Staubli VAL3: HMI_safezone.pjx

--- HMI_safezone.pjx ---
Parameters version=s8.15Cs9_BS3113 stackSize=5000 millimeterUnit=true
Program file=bind.pgx
Program file=main.pgx
Program file=movePoint.pgx
Program file=onStart.pgx
Program file=refreshData.pgx
Program file=setData.pgx
Program file=setFrameData.pgx
Program file=start.pgx
Program file=stop.pgx
Program file=teachPoint.pgx
Data file=HMI_safezone.dtx
Library alias=safeTemp path=Disk://data/CustomerLib/default/safeData/safeData.pjx
Library alias=util path=Disk://HMI_cs9/HMI_util/HMI_util.pjx
Library alias=safeCheck path=Disk://source/projectSource/safeCheck/safeCheck.pjx
Library alias=saveData path=Disk://source/saveData/saveData.pjx

--- HMI_safezone.dtx ---
mdesc mNomSpeed = {blend=off}
string sList
string sSelZone
bool bSetFrame
bool bTeach1
bool bMove
bool bRename
bool bConfirm
bool bActive
public num nFrame[6]
num nTRSF1[6]
num nTRSF2[6]
string sLastZone
num _nZoneIndex
string sComment
frame fFrame = {fatherId=world[0]}
bool bBack
tool tTool = {fatherId=flange[0]}
bool bSetFrameData
string sToolIndex

--- main.pgx ---
public program main()
  local bool l_bResult
  local bool l_bExit
begin
  do
    if util:sPage!="safezone"
      util:sPage="safezone"
      call util:loadingPage()
      call onStart()
      call bind()
      userPage(util:sPage)
      delay(0.5)
    endIf

    if sSelZone!=sLastZone and sSelZone!=""
      sLastZone=sSelZone
      toNum(sLastZone,_nZoneIndex,l_bResult)
      bActive=(safeTemp:zZoneItem[_nZoneIndex].bActive==true)
      call refreshData(_nZoneIndex)
    endIf
    if bSetFrame
      //      util:sPage="Wizard"
      //      userPage(util:sPage)
      bSetFrame=false
      //      popUpMsg("设定坐标系")
      //      call refreshData(_nZoneIndex)
    elseIf bSetFrameData
      bSetFrameData=false
      call setFrameData(_nZoneIndex)
      call refreshData(_nZoneIndex)

    elseIf bTeach1
      bTeach1=false
      call teachPoint(_nZoneIndex)
      call refreshData(_nZoneIndex)
    elseIf bMove
      bMove=false
      call movePoint(_nZoneIndex)
    elseIf bConfirm
      bConfirm=false
      call setData(_nZoneIndex)
      call refreshData(_nZoneIndex)
    elseIf bBack
      bBack=false
      l_bExit=true
    endIf

    delay(0)
  until l_bExit==true
  call saveData:setBaseJOG(saveData:nJogTool)
end

--- start.pgx ---
program start()
begin
end

--- bind.pgx ---
program bind()
  local string l_nmb
  local num l_i
begin
  userPageBindClick("safezone","btnback",bBack,true)
  //
  userPageBind("safezone","cbx1","options",sList,size(sList),"r")
  userPageBind("safezone","cbx1","value",sSelZone,1,"rw")

  userPageBindClick("safezone","btn1",bSetFrame,true)
  userPageBindClick("safezone","btn2",bTeach1,true)
  userPageBindClick("safezone","btn2_Copy1",bMove,true)
  // userPageBindClick("safezone","btn3",bRename,true)
  userPageBindClick("safezone","btn4",bConfirm,true)
  userPageBindClick("safezone","btnSetFrame",bSetFrameData,true)

  userPageBind("safezone","txt1","value",sComment,1,"rw")

  userPageBind("safezone","chk1","checked",bActive,1,"rw")

  //  userPageBindClick("Wizard","btn1",bExit,true)


  for l_i = 0 to 5
    l_nmb="nmb"+toString("",l_i)
    userPageBind("safezone",l_nmb,"value",nFrame[l_i],1,"rw")
  endFor

  for l_i = 0 to 5
    l_nmb="nmb1"+toString("",l_i)
    userPageBind("safezone",l_nmb,"value",nTRSF1[l_i],1,"rw")
  endFor

  for l_i = 0 to 5
    l_nmb="nmb2"+toString("",l_i)
    userPageBind("safezone",l_nmb,"value",nTRSF2[l_i],1,"rw")
  endFor
end

--- movePoint.pgx ---
public program movePoint(num x_nIndex)
  local pointRx l_pPoint
  local bool l_bResult
  local tool l_tTool
begin

  l_bResult=userPageConfirm("是否移动到此点位？")

  if l_bResult
    resetMotion()
    link(l_pPoint,fFrame)
    call saveData:getTool(saveData:nJogTool,l_tTool)
    l_pPoint.trsf=safeTemp:zZoneItem[x_nIndex].pFirst.trsf
    l_pPoint.config=safeTemp:zZoneItem[x_nIndex].pFirst.config
    movej(l_pPoint,l_tTool,mNomSpeed)
    delay(0)
  endIf
end

--- onStart.pgx ---
program onStart()
  local num l_i
  local num l_nResult
begin
  call saveData:setBaseJOG(saveData:nJogTool)
  sToolIndex=toString("",saveData:nJogTool)
  sSelZone=""
  sLastZone=""
  resize(sList,1,size(safeTemp:zZoneItem))

  for l_i = 0 to size(sList)-1
    sList[l_i]=toString("",l_i)+","+safeTemp:zZoneItem[l_i].sID
  endFor
  bActive=false
  for l_i = 0 to 5
    nFrame[l_i]=0
    nTRSF1[l_i]=0
    nTRSF2[l_i]=0
  endFor
end

--- refreshData.pgx ---
program refreshData(num x_nIndex)
  local tool l_tTool
begin
  nFrame[0]=safeTemp:zZoneItem[x_nIndex].fBase.trsf.x
  nFrame[1]=safeTemp:zZoneItem[x_nIndex].fBase.trsf.y
  nFrame[2]=safeTemp:zZoneItem[x_nIndex].fBase.trsf.z
  nFrame[3]=safeTemp:zZoneItem[x_nIndex].fBase.trsf.rx
  nFrame[4]=safeTemp:zZoneItem[x_nIndex].fBase.trsf.ry
  nFrame[5]=safeTemp:zZoneItem[x_nIndex].fBase.trsf.rz
  fFrame.trsf=safeTemp:zZoneItem[x_nIndex].fBase.trsf
  call saveData:getTool(saveData:nJogTool,tTool)
  $jogContext(tTool,fFrame,0)

  nTRSF1[0]=safeTemp:zZoneItem[x_nIndex].pFirst.trsf.x
  nTRSF1[1]=safeTemp:zZoneItem[x_nIndex].pFirst.trsf.y
  nTRSF1[2]=safeTemp:zZoneItem[x_nIndex].pFirst.trsf.z
  nTRSF1[3]=safeTemp:zZoneItem[x_nIndex].pFirst.trsf.rx
  nTRSF1[4]=safeTemp:zZoneItem[x_nIndex].pFirst.trsf.ry
  nTRSF1[5]=safeTemp:zZoneItem[x_nIndex].pFirst.trsf.rz

  nTRSF2[0]=safeTemp:zZoneItem[x_nIndex].pSecond.trsf.x
  nTRSF2[1]=safeTemp:zZoneItem[x_nIndex].pSecond.trsf.y
  nTRSF2[2]=safeTemp:zZoneItem[x_nIndex].pSecond.trsf.z
  nTRSF2[3]=safeTemp:zZoneItem[x_nIndex].pSecond.trsf.rx
  nTRSF2[4]=safeTemp:zZoneItem[x_nIndex].pSecond.trsf.ry
  nTRSF2[5]=safeTemp:zZoneItem[x_nIndex].pSecond.trsf.rz

  sComment=safeTemp:zZoneItem[x_nIndex].sID

end

--- setData.pgx ---
public program setData(num x_nIndex)
  local pointRx l_pPoint
begin
  safeTemp:zZoneItem[x_nIndex].fBase.trsf.x=nFrame[0]
  safeTemp:zZoneItem[x_nIndex].fBase.trsf.y=nFrame[1]
  safeTemp:zZoneItem[x_nIndex].fBase.trsf.z=nFrame[2]
  safeTemp:zZoneItem[x_nIndex].fBase.trsf.rx=nFrame[3]
  safeTemp:zZoneItem[x_nIndex].fBase.trsf.ry=nFrame[4]
  safeTemp:zZoneItem[x_nIndex].fBase.trsf.rz=nFrame[5]


  safeTemp:zZoneItem[x_nIndex].pFirst.trsf.x=nTRSF1[0]
  safeTemp:zZoneItem[x_nIndex].pFirst.trsf.y=nTRSF1[1]
  safeTemp:zZoneItem[x_nIndex].pFirst.trsf.z=nTRSF1[2]
  safeTemp:zZoneItem[x_nIndex].pFirst.trsf.rx=nTRSF1[3]
  safeTemp:zZoneItem[x_nIndex].pFirst.trsf.ry=nTRSF1[4]
  safeTemp:zZoneItem[x_nIndex].pFirst.trsf.rz=nTRSF1[5]

  safeTemp:zZoneItem[x_nIndex].pSecond.trsf.x=nTRSF2[0]
  safeTemp:zZoneItem[x_nIndex].pSecond.trsf.y=nTRSF2[1]
  safeTemp:zZoneItem[x_nIndex].pSecond.trsf.z=nTRSF2[2]
  safeTemp:zZoneItem[x_nIndex].pSecond.trsf.rx=nTRSF2[3]
  safeTemp:zZoneItem[x_nIndex].pSecond.trsf.ry=nTRSF2[4]
  safeTemp:zZoneItem[x_nIndex].pSecond.trsf.rz=nTRSF2[5]



  safeTemp:zZoneItem[x_nIndex].bActive=(bActive==true)
  safeTemp:zZoneItem[x_nIndex].sID=sComment

  safeTemp:libSave()
  delay(0.1)
  popUpMsg("safedata已保存")

end

--- setFrameData.pgx ---
program setFrameData(num x_nIndex)
  local bool l_bResult
  local num l_nResult
begin

  l_bResult=userPageConfirm("确定设定坐标系？(点位会随坐标系改变)")

  if l_bResult
    safeTemp:zZoneItem[x_nIndex].fBase.trsf.x=nFrame[0]
    safeTemp:zZoneItem[x_nIndex].fBase.trsf.y=nFrame[1]
    safeTemp:zZoneItem[x_nIndex].fBase.trsf.z=nFrame[2]
    safeTemp:zZoneItem[x_nIndex].fBase.trsf.rx=nFrame[3]
    safeTemp:zZoneItem[x_nIndex].fBase.trsf.ry=nFrame[4]
    safeTemp:zZoneItem[x_nIndex].fBase.trsf.rz=nFrame[5]
    fFrame.trsf=safeTemp:zZoneItem[x_nIndex].fBase.trsf

    l_nResult=safeTemp:libSave()
    if l_nResult==0
      popUpMsg("设定坐标系完成")
    else
      popUpMsg("设定坐标系失败")
    endIf
  endIf
end

--- stop.pgx ---
program stop()
begin
end

--- teachPoint.pgx ---
program teachPoint(num x_nIndex)
  local bool l_bResult
  local pointRx l_pPoint
  local tool l_tTool
begin
  l_bResult=userPageConfirm("是否记录当前点位？")
  if l_bResult
    call saveData:getTool(saveData:nJogTool,l_tTool)
    fFrame.trsf.x=nFrame[0]
    fFrame.trsf.y=nFrame[1]
    fFrame.trsf.z=nFrame[2]
    fFrame.trsf.rx=nFrame[3]
    fFrame.trsf.ry=nFrame[4]
    fFrame.trsf.rz=nFrame[5]

    l_pPoint=here(l_tTool,fFrame)
    safeTemp:zZoneItem[x_nIndex].pFirst.trsf=l_pPoint.trsf
    safeTemp:zZoneItem[x_nIndex].pFirst.config=l_pPoint.config
    safeTemp:libSave()




    delay(0.1)
  endIf
end
